Fanuc KAREL source: KD00050.KL

PROGRAM KD00050
%NOLOCKGROUP
%DEFGROUP = 1
VAR
  I: INTEGER
  J: INTEGER
  B: BOOLEAN
  R: REAL
  S: STRING[80]
BEGIN
  MOVE AXIS 1 BY 10.0
END KD00050
